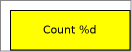
VISUALIZATION VisuB1x  // 132x52
    Rectangle (10,10 120x40), "Count %d", tooltip "rect tip", text variable: GVL_Fixture.nCount, invisible if: GVL_Fixture.bEnable, input disabled if: NOT GVL_Fixture.bEnable
        p3560616238: GVL_Fixture.nCount
        p2738717112: GVL_Fixture.nCount
        p2858320360: GVL_Fixture.nCount
END_VISUALIZATION

(* stored: Version 1.1.0.1
   Visu VisuB1x: Id {7762283b-ef9c-4e21-bd1f-25399c002855} *)
